Fanuc KAREL source: kx00008.KL

-- PROVISIONAL review KL for V1013-1; original PC SHA256 75304a9b45cb0f1e2c7d29907f6d69c8bca444b36d217644031e4f1fb12085bb
-- Incomplete behavior may be omitted. Consult companion uncertainty JSON. Do not deploy.
PROGRAM KX00008
%NOLOCKGROUP
VAR
  I : INTEGER
  J : INTEGER
  B : BOOLEAN
  F : FILE
  S : STRING[80]
-- UNRESOLVED_DECL P type=000102
BEGIN
  -- UNRESOLVED_PC offsets 5-7; opcodes 9C,3A
  -- UNRESOLVED_PC offsets 12-16; opcodes 7F
END KX00008
